(* IEC 61131-3 sources: 2026_Projet_YGO_ExcavatriceDragage/CODE_BACKUP/CODE_20260904_AvantWeekendBackup_v0.6.34/B_AU_SECURITE/_TYPES, 4 files *)

(* ---- ST_Safety_Emergency_Cmd.st ---- *)
(* =======================================================================
   ⚙️ ST_Safety_Emergency_Cmd — Commandes de pilotage de la chaîne AU
   ───────────────────────────────────────────────────────────────
   🎯 Rôle : DUT de commande du FB_Safety_EmergencyManagement fusionné.
      Regroupe les commandes physiques fail-safe de pilotage des canaux
      de maintien et de l'impulsion de réarmement.
   🔒 Polarité : MaintainA/B_Cmd en maintien (TRUE = voie saine).
      Fail-safe : Enable=FALSE → toutes commandes à FALSE.
   🔌 Interface : Produit par FB_Safety_EmergencyManagement.Cmd, consommé par
      PRG_06_Outputs uniquement.
   📄 Doc métier : DOC/AF/AF_Partie-01_Analyse_Fonctionnelle_v2.1.md
   ======================================================================= *)

TYPE ST_Safety_Emergency_Cmd :
STRUCT
    MaintainA_Cmd   : BOOL; // <-- [ACT]  Sortie pilotage canal A (TRUE = voie maintenue)
    MaintainB_Cmd   : BOOL; // <-- [ACT]  Sortie pilotage canal B (TRUE = voie maintenue)
    ArmPulse_Cmd    : BOOL; // <-- [ACT]  Impulsion rearmement physique (1s)
    TestCutActive   : BOOL; // <-- [ACT]  Test de redondance en cours (canal A ou B coupe) — consommé par la simulation
END_STRUCT
END_TYPE

(* ---- ST_Safety_Emergency_Diag.st ---- *)
(* =======================================================================
   📊 ST_Safety_Emergency_Diag — Diagnostic et erreurs de la chaîne AU
   ───────────────────────────────────────────────────────────────
   🎯 Rôle : Structure de diagnostic et erreurs de la chaîne d'arrêt d'urgence
   🔌 Interface : Produit par FB_Safety_EmergencyManagement, consommé par Supervision/Troubleshooting
   📄 Doc métier : DOC/AF/AF_Partie-01_Analyse_Fonctionnelle_v2.1.md
   ======================================================================= *)

TYPE ST_Safety_Emergency_Diag :
STRUCT
    Error                : BOOL; // Synthese defaut active : (ErrorId <> 0)
    ErrorId              : WORD; // Bitfield erreurs : bit0=Redundancy, bit1=Arming, bit3=Startup
    RedundancyTestFailed : BOOL; // Canal A ou B reste colle/shunte detecte a l'auto-test (Reset requis)
    ArmFailed            : BOOL; // Impulsion envoyee mais contacteur puissance non confirme sous 2s (Reset requis)
    WasArmed             : BOOL; // TRUE = AU armee au moins une fois (contacteur confirme) ; maintien PowerKeepAlive a travers un appui AU pur — retombe sur raison metier (coupure/redondance/Enable OFF)
    LockoutActive        : BOOL; // Verrouillage temporel de 5s entre tentatives de rearmement echouees
    LastAbortStep        : INT;  // Etape de la sequence AU lors du dernier abandon (0 a 6)
    LastAbortCause       : WORD; // Bitfield cause abandon : 16#0001=Cut IHM, 16#0002=Chute chaine pulse/confirm, 16#0004=Timeout A, 16#0008=Timeout B, 16#0010=PowerCutOff metier
END_STRUCT
END_TYPE

(* ---- ST_Safety_Emergency_State.st ---- *)
(* =======================================================================
   📊 ST_Safety_Emergency_State — État public de la chaîne d'arrêt d'urgence
   ───────────────────────────────────────────────────────────────
   🎯 Rôle : Bus d'état public de la chaîne d'arrêt d'urgence
   🔌 Interface : Produit par FB_Safety_EmergencyManagement, consommé par Supervision/Troubleshooting
   📄 Doc métier : DOC/AF/AF_Partie-01_Analyse_Fonctionnelle_v2.1.md
   ======================================================================= *)

TYPE ST_Safety_Emergency_State :
STRUCT
    ChainOk     : BOOL; // Boucle AU fermee (EmergencyChainClosed = TRUE)
    ContactorOk : BOOL; // Contacteur puissance confirme engage (PowerContactorEngaged = TRUE)
    Step        : INT;  // Etape sequence armement : 0=IDLE, 1=TestA, 2=RestoreA, 3=TestB, 4=RestoreB, 5=Pulse, 6=Confirm
    Armable     : BOOL; // Rearmement possible maintenant : chain OK, step=0, pas de lockout
    ArmingBusy  : BOOL; // Sequence armement OU lockout en cours (nouvelle demande ignoree)
END_STRUCT
END_TYPE

(* ---- ST_Safety_Emergency_Status.st ---- *)
(* =======================================================================
   📊 ST_Safety_Emergency_Status — État & diagnostic de la chaîne AU
   ───────────────────────────────────────────────────────────────
   🎯 Rôle : DUT d'état/diagnostic du FB_Safety_EmergencyManagement fusionné.
      Regroupe les états publics IEC (Ready/Done), le bus d'état (State),
      le bus de diagnostic (Diag), le défaut laté (Fault : ST_Fault, socle
      FB_FaultCore) et le message opérateur par état / par problème.
   🔒 Sécurité : interlock TOUJOURS sur la cause brute (State/Diag), jamais sur le latch.
      Fail-safe : Enable=FALSE → Ready à FALSE.
   🔌 Interface : Produit par FB_Safety_EmergencyManagement.Status, consommé par
      PRG_07_Supervision / IHM / Troubleshooting.
   📄 Doc métier : DOC/AF/AF_Partie-01_Analyse_Fonctionnelle_v2.1.md
   ======================================================================= *)

TYPE ST_Safety_Emergency_Status :
STRUCT
    // === ETATS PUBLICS IEC ===
    Ready           : BOOL; // <-- [STAT] FB pret a fonctionner (Enable + pas de StartupFail)
    Done            : BOOL; // <-- [STAT] Contacteur puissance confirme engage

    // === BUS D'ETAT & DIAGNOSTIC ===
    State           : ST_Safety_Emergency_State; // <-- [STAT] Bus d'etat public
    Diag            : ST_Safety_Emergency_Diag;  // <-- [DIAG] Bus de diagnostic public

    // === DEFAUT LATCHE (socle FB_FaultCore) ===
    Fault           : ST_Fault; // <-- [DIAG] Brique defaut (vue live + latchee), corrige le bug bit3 StartupFail

    // === MESSAGE OPERATEUR PAR ETAT / PAR PROBLEME ===
    OperatorMessage : STRING(120); // <-- [DIAG] Message explicite par etat / par probleme de la chaine AU
END_STRUCT
END_TYPE
